Fanuc KAREL source: kt00523.KL

-- PROVISIONAL review KL for V940-1; original PC SHA256 8f1aff95fd52bfc5aa8d18a479711138bd13ae5b608ac52683cc08c324d24957
-- Incomplete behavior may be omitted. Consult companion uncertainty JSON. Do not deploy.
PROGRAM KT00523
%NOLOCKGROUP
VAR
  OUT : BOOLEAN
-- UNRESOLVED_DECL P1 type=000106
-- UNRESOLVED_DECL P2 type=000106
BEGIN
  -- V9_ZERO_TABLE_METADATA_HINT layout=0001; no indexed target words; source/name/runtime held
  -- UNRESOLVED_PC offsets 5-20; opcodes 2E,22,32,35
  -- UNRESOLVED_PC offsets 25-40; opcodes 2E,22,32,35
  -- UNRESOLVED_PC offsets 45-60; opcodes 2E,22,32,35
  -- UNRESOLVED_PC offsets 65-80; opcodes 2E,22,32,35
  -- UNRESOLVED_PC offsets 85-118; opcodes 49,7E,49,7E,AC,23
  -- UNRESOLVED_PC offsets 123-127; opcodes 7F
END KT00523
